Fanuc KAREL source: ko00108.KL

-- PROVISIONAL review KL for V940-1; original PC SHA256 835b92d3fceb5da5cee654deb9cbe47e4b50a65bf95e9f4cc80f496283e49eaa
-- Incomplete behavior may be omitted. Consult companion uncertainty JSON. Do not deploy.
PROGRAM KO00108
%NOLOCKGROUP
VAR
  A : REAL
  B : REAL
  OUT : REAL
BEGIN
  -- V9_ZERO_TABLE_METADATA_HINT layout=0001; no indexed target words; source/name/runtime held
  -- UNRESOLVED_PC offsets 5-13; opcodes 9D,64,23
  -- UNRESOLVED_PC offsets 18-30; opcodes 2E,64,23
  -- UNRESOLVED_PC offsets 35-56; opcodes 27,22,22,76,23
  -- UNRESOLVED_PC offsets 61-65; opcodes 7F
END KO00108
